Universal Robots PolyScope program: TurnProg.urp

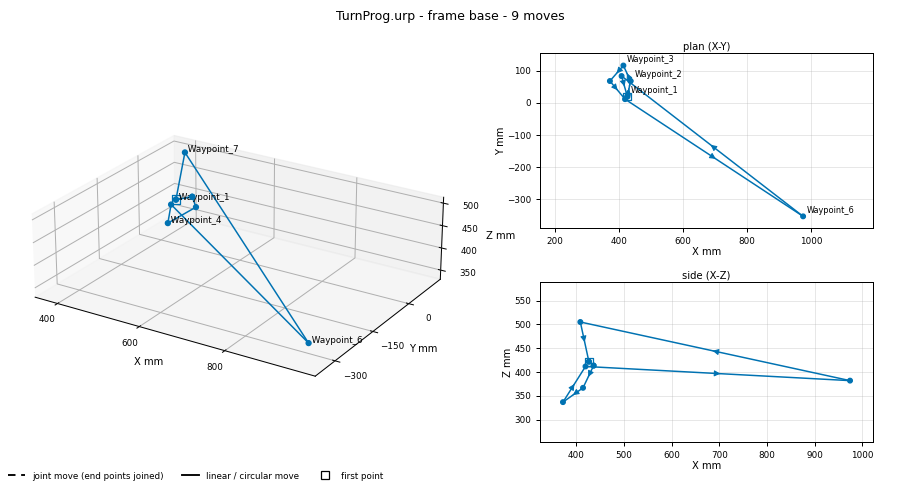
[picture p0: tool path of TurnProg.urp in frame base, 9 of 9 moves have a stored position in this frame; points joined in program order, loops and branches not executed]
Program TurnProg (createdIn=3.0.0 lastSavedIn=3.0.0 directory=/programs installation=default)
Robot Program (runOnlyOnce=true motionType=MoveJ speed=1.047198 acceleration=1.396263 useActiveTCP=false)
  'Program generated by RoboDK v6.0.7 for ABB IRB 120-3/0.6 on XX/XX/XXXX 18:00:00'
  'Using nominal kinematics.'
  'Using Ref. Frame S: p[1.234570, -0.098765, 0.050500, 0.000000, 0.000000, 0.523599]'
  'Using TCP Tool S: p[0.010000, 0.020000, 0.150000, 0.000000, 0.000000, 0.000000]'
  Script: set_tcp(p[0.010000, 0.020000, 0.150000, 0.000000, 0.000000, 0.000000])
  MoveL speed 250 mm/s, acceleration 1200 mm/s^2 (useActiveTCP=true)
    Waypoint Waypoint_1: TCP in base x=426.318 y=20 z=422.034 mm, rx=0.1383 ry=2.2532 rz=-0.2966 rad; joints [200, 0, 0, 0, 30, 0] deg; flange x=317.789 y=39.504 z=526.155 mm, rx=0.1383 ry=2.2532 rz=-0.2966 rad
    Waypoint Waypoint_2: TCP in base x=436.232 y=68.297 z=413.715 mm, rx=0.1383 ry=2.2532 rz=-0.2966 rad; joints [0, 0, 0, -200, 30, 0] deg; flange x=327.703 y=87.801 z=517.836 mm, rx=0.1383 ry=2.2532 rz=-0.2966 rad
    Waypoint Waypoint_3: TCP in base x=414.005 y=116.593 z=367.095 mm, rx=0.1383 ry=2.2532 rz=-0.2966 rad; joints [0, 0, 0, 0, 30, 200] deg; flange x=305.476 y=136.097 z=471.216 mm, rx=0.1383 ry=2.2532 rz=-0.2966 rad
    Waypoint Waypoint_4: TCP in base x=371.953 y=68.296 z=337.111 mm, rx=0.1383 ry=2.2532 rz=-0.2966 rad; joints [-200, 0, 0, 0, 30, -200] deg; flange x=263.425 y=87.801 z=441.232 mm, rx=0.1383 ry=2.2532 rz=-0.2966 rad
    Waypoint Waypoint_5: TCP in base x=419.189 y=11.793 z=411.899 mm, rx=0.1383 ry=2.2532 rz=-0.2966 rad; joints [0, 190, -190, 0, 190, 0] deg; flange x=310.661 y=31.298 z=516.02 mm, rx=0.1383 ry=2.2532 rz=-0.2966 rad
    Waypoint Waypoint_6: TCP in base x=973.908 y=-353.337 z=382.202 mm, rx=-0.5037 ry=2.3595 rz=0.0001 rad; joints [-90, -30, 60, 180, -30, -180] deg; flange x=890.027 y=-389.125 z=503.376 mm, rx=-0.5037 ry=2.3595 rz=0.0001 rad
    Waypoint Waypoint_7: TCP in base x=408.367 y=83.8 z=505.12 mm, rx=-0.4874 ry=1.4458 rz=-0.7473 rad; joints [350, 0, 0, -350, 30, 540] deg; flange x=257.546 y=97.782 z=512.713 mm, rx=-0.4874 ry=1.4458 rz=-0.7473 rad
    Waypoint Waypoint_8: TCP in base x=426.318 y=20 z=422.034 mm, rx=0.1383 ry=2.2532 rz=-0.2966 rad; joints [-180, 0, 0, 180, 0, -540] deg; flange x=317.789 y=39.504 z=526.155 mm, rx=0.1383 ry=2.2532 rz=-0.2966 rad
  Script: movej([6.108652, 0.000000, 0.000000, -6.108652, 0.523599, 9.424778],1.20000,0.75000,0,0.0000)
  MoveJ speed 42.97 deg/s, acceleration 68.75 deg/s^2 (useActiveTCP=true)
    Waypoint Waypoint_9: TCP in base x=436.232 y=68.297 z=413.715 mm, rx=0.1383 ry=2.2532 rz=-0.2966 rad; joints [350, 0, 0, -350, 30, 540] deg; flange x=327.703 y=87.801 z=517.836 mm, rx=0.1383 ry=2.2532 rz=-0.2966 rad
